(* Logix 5000 project; controller R400_500_XLS vendor 1 type 14 code 216 rev 31.11; software revision 31.01; part 31 of 32 *)
(* tags used below, declared in another part *)
   Abort1 : DINT;   // Not Used
   CycExcBuffer : UDT_CYCLE;
   CycleSequence : UDT_CYCLE_SEQUENCE;
   DintBuffer : DINT[5];
   DRYING : DINT;   // Drying id number
   M : DINT[5];   // Memory Bits
   OneShot : DINT[1];
   ONS_FC64 : DINT;
   PREWASH_1 : DINT;   // Pre-wash 1 id number
   PREWASH_2 : DINT;   // Pre-wash 2 id number
   PREWASH_3 : DINT;   // Pre-wash 3 id number
   PREWASH_4 : DINT;   // Pre-wash 4 id number
   PwExcBuffer : UDT_PW;
   PWR_UP : DINT;
   rBuffer : REAL[4];
   rIn_WSH61 : REAL;
   RINSE_1 : DINT;   // Rinse 1 id number
   RINSE_2 : DINT;   // Rinse 2 id number
   RINSE_3 : DINT;   // Rinse 3 id number
   RinseExcBuffer : UDT_RINSE;
   Run : DINT;
   sOut_WSH61 : STRING;
   String : STRING[50];   // String
   Tmr : TIMER[107];
   WASH_1 : DINT;   // Wash 1 id number
   WASH_2 : DINT;   // Wash 2 id number
   WASH_3 : DINT;   // Wash 3 id number
   WASH_4 : DINT;   // Wash 4 id number
   WASH_5 : DINT;   // Wash 5 id number
   WshExcBuffer : UDT_WASH;
   ActualDay : DINT;
   Current_Screen : DINT;
   DateTime : DINT[7];
   Doors_Check : DINT;
   DoorSafetyCheck : BOOL;
   DoorSafetyCheckDay : DINT;
   DoorSafetyCheckMonth : DINT;
   DoorSafetyCheckYear : DINT;
   I_Ld_Dr_Cls_Sw : BOOL;   // Load door close
   I_Ld_Dr_Obs_Sw : BOOL;   // Load door obstruction switch
   I_Unld_Dr_Cls_Sw : BOOL;   // Unload door close
   I_Unld_Dr_Obs_Sw : BOOL;   // Unload door obstruction switch
   LastCheckNbrDays : DINT;
   Load : Doors;
   MaintainCloseLd : BOOL;
   MaintainCloseUnld : BOOL;
   MaintainOpenLd : BOOL;
   MaintainOpenUnld : BOOL;
   MaintenanceDueDays : DINT;
   msg : BOOL[512];
   Msg_DoorSteps : INT;   // Display Safety Door Test Messages
   ONS_WSH64 : SINT;
   RecallSafetyCheck : BOOL;
   Screen_Ctrl : DINT;   // PLC Screen Request
   Tpb : DINT[11];
   TpbImage : DINT[11];
   TreatmentPtr : DINT;
   Unit : Hrdwre;   // Unit Configuration
   UnLoad : Doors;
(* MainProgram, continued *)

ROUTINE WSH_61_Real_to_String   (* ladder *)
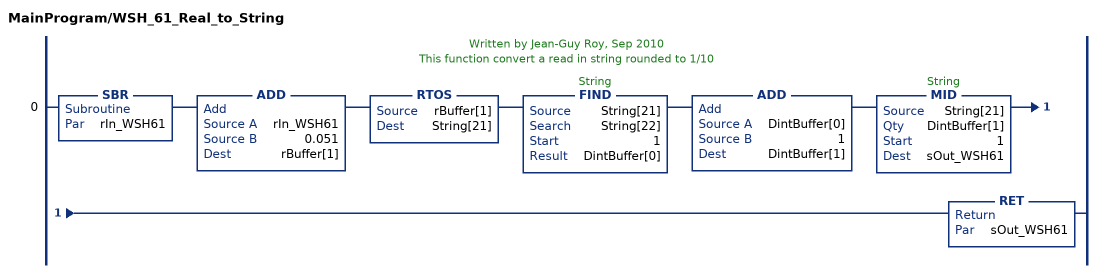
   // Written by Jean-Guy Roy, Sep 2010
   // This function convert a read in string rounded to 1/10
   0: SBR(rIn_WSH61)ADD(rIn_WSH61,0.051,rBuffer[1])RTOS(rBuffer[1],String[21])FIND(String[21],String[22],1,DintBuffer[0])ADD(DintBuffer[0],1,DintBuffer[1])MID(String[21],DintBuffer[1],1,sOut_WSH61)RET(sOut_WSH61);
END_ROUTINE

ROUTINE WSH_64_DOOR_MAINTENANCE   (* ladder *)
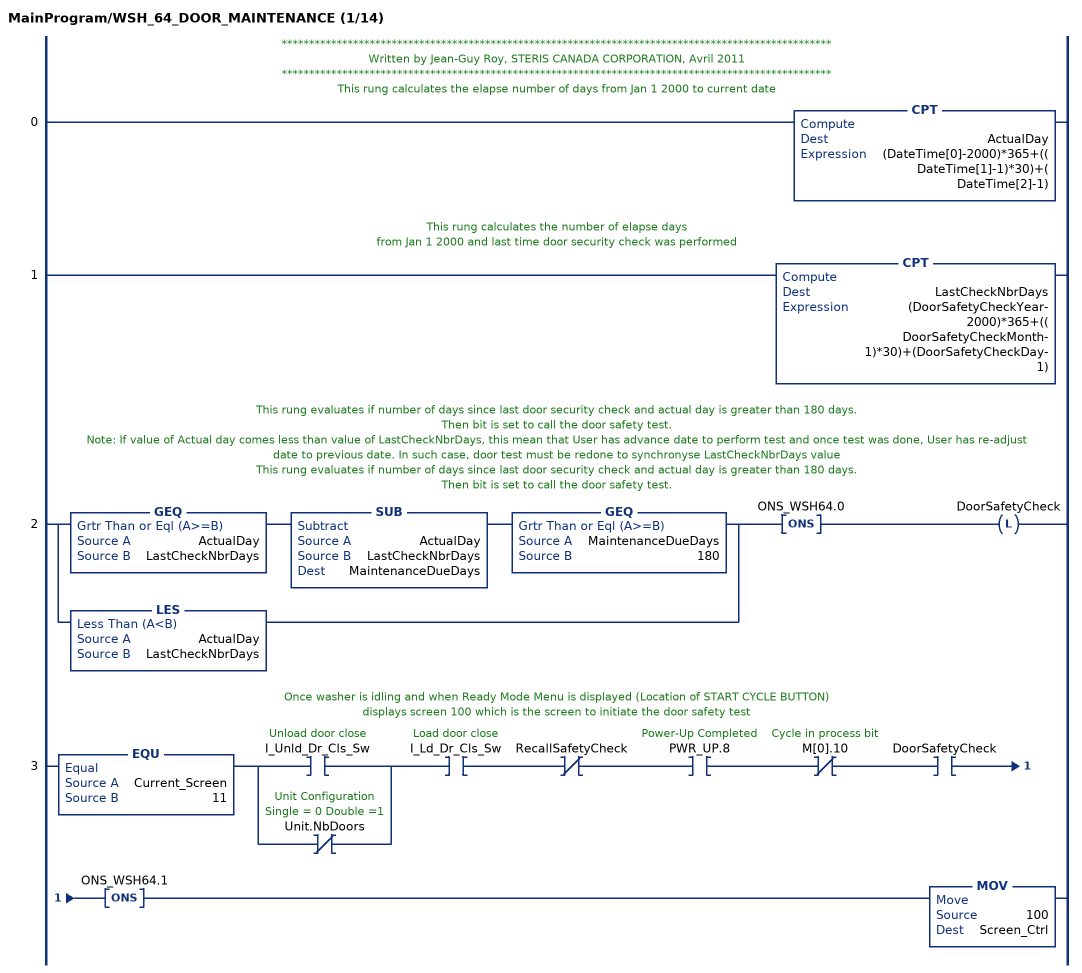
   // ****************************************************************************************************
   // Written by Jean-Guy Roy, STERIS CANADA CORPORATION, Avril 2011
   // ****************************************************************************************************
   // This rung calculates the elapse number of days from Jan 1 2000 to current date
   0: CPT(ActualDay,(DateTime[0]-2000)*365+((DateTime[1]-1)*30)+(DateTime[2]-1));
   // This rung calculates the number of elapse days
   // from Jan 1 2000 and last time door security check was performed
   1: CPT(LastCheckNbrDays,(DoorSafetyCheckYear-2000)*365+((DoorSafetyCheckMonth-1)*30)+(DoorSafetyCheckDay-1));
   // This rung evaluates if number of days since last door security check and actual day is greater than 180 days.
   // Then bit is set to call the door safety test.
   // Note: If value of Actual day comes less than value of LastCheckNbrDays, this mean that User has advance date to perform test and once test was done, User has re-adjust date to previous date. In such case, door test must be redone to synchronyse LastCheckNbrDays value
   // This rung evaluates if number of days since last door security check and actual day is greater than 180 days.
   // Then bit is set to call the door safety test.
   2: [GEQ(ActualDay,LastCheckNbrDays) SUB(ActualDay,LastCheckNbrDays,MaintenanceDueDays) GEQ(MaintenanceDueDays,180) ,LES(ActualDay,LastCheckNbrDays) ]ONS(ONS_WSH64.0)OTL(DoorSafetyCheck);
   // Once washer is idling and when Ready Mode Menu is displayed (Location of START CYCLE BUTTON)
   // displays screen 100 which is the screen to initiate the door safety test
   3: EQU(Current_Screen,11)[XIC(I_Unld_Dr_Cls_Sw) ,XIO(Unit.NbDoors) ]XIC(I_Ld_Dr_Cls_Sw)XIO(RecallSafetyCheck)XIC(PWR_UP.8)XIO(M[0].10)XIC(DoorSafetyCheck)ONS(ONS_WSH64.1)MOV(100,Screen_Ctrl);
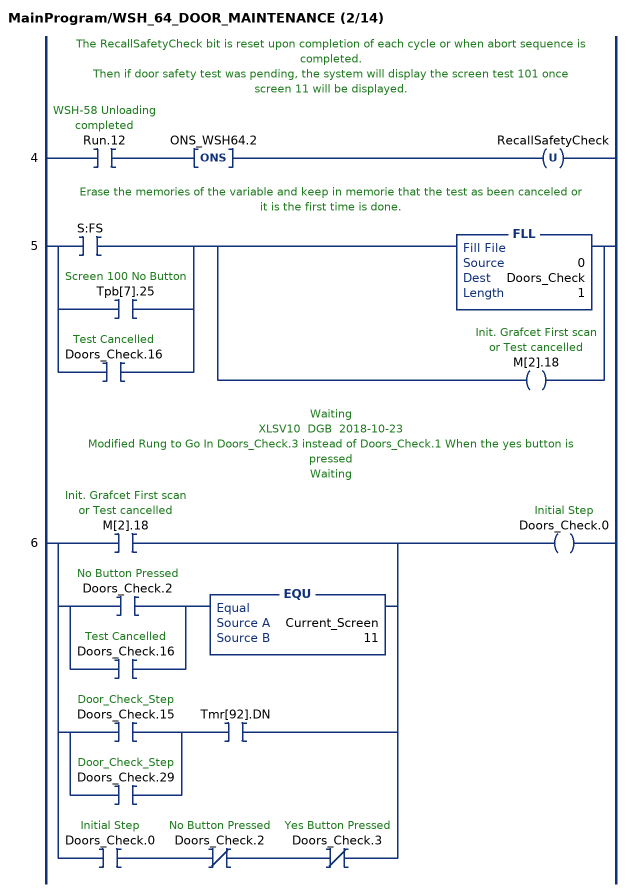
   // The RecallSafetyCheck bit is reset upon completion of each cycle or when abort sequence is completed.
   // Then if door safety test was pending, the system will display the screen test 101 once screen 11 will be displayed.
   4: XIC(Run.12)ONS(ONS_WSH64.2)OTU(RecallSafetyCheck);
   // Erase the memories of the variable and keep in memorie that the test as been canceled or it is the first time is done.
   5: [XIC(S:FS) ,XIC(Tpb[7].25) ,XIC(Doors_Check.16) ][FLL(0,Doors_Check,1) ,OTE(M[2].18) ];
   // Waiting
   // XLSV10  DGB  2018-10-23
   // Modified Rung to Go In Doors_Check.3 instead of Doors_Check.1 When the yes button is pressed
   // Waiting
   6: [XIC(M[2].18) ,[XIC(Doors_Check.2) ,XIC(Doors_Check.16) ] EQU(Current_Screen,11) ,[XIC(Doors_Check.15) ,XIC(Doors_Check.29) ] XIC(Tmr[92].DN) ,XIC(Doors_Check.0) XIO(Doors_Check.2) XIO(Doors_Check.3) ]OTE(Doors_Check.0);
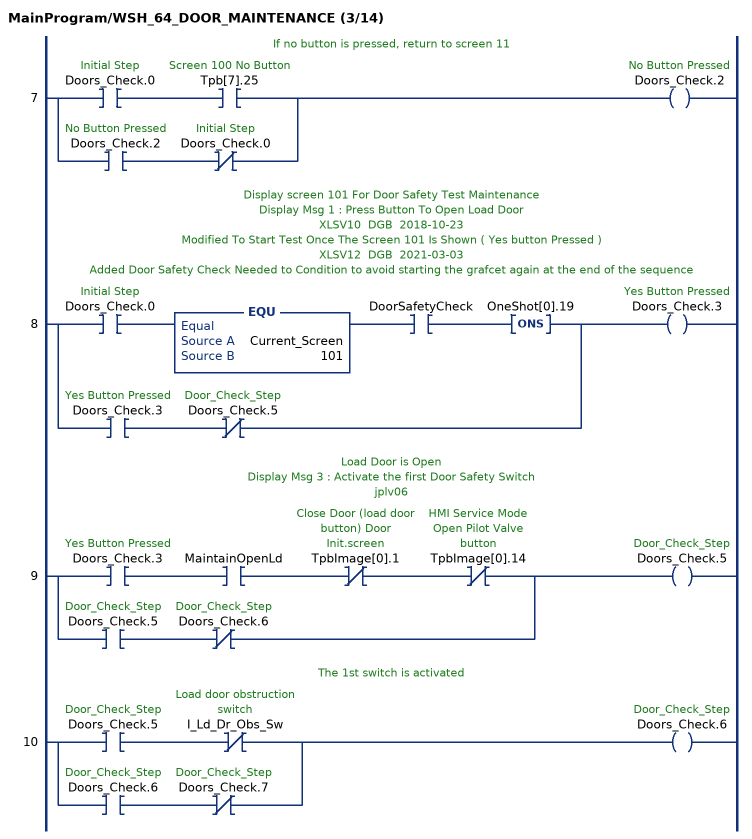
   // If no button is pressed, return to screen 11
   7: [XIC(Doors_Check.0) XIC(Tpb[7].25) ,XIC(Doors_Check.2) XIO(Doors_Check.0) ]OTE(Doors_Check.2);
   // Display screen 101 For Door Safety Test Maintenance
   // Display Msg 1 : Press Button To Open Load Door
   // XLSV10  DGB  2018-10-23
   // Modified To Start Test Once The Screen 101 Is Shown ( Yes button Pressed )
   // XLSV12  DGB  2021-03-03
   // Added Door Safety Check Needed to Condition to avoid starting the grafcet again at the end of the sequence
   8: [XIC(Doors_Check.0) EQU(Current_Screen,101) XIC(DoorSafetyCheck) ONS(OneShot[0].19) ,XIC(Doors_Check.3) XIO(Doors_Check.5) ]OTE(Doors_Check.3);
   // Load Door is Open
   // Display Msg 3 : Activate the first Door Safety Switch
   // jplv06
   9: [XIC(Doors_Check.3) XIC(MaintainOpenLd) XIO(TpbImage[0].1) XIO(TpbImage[0].14) ,XIC(Doors_Check.5) XIO(Doors_Check.6) ]OTE(Doors_Check.5);
   // The 1st switch is activated
   10: [XIC(Doors_Check.5) XIO(I_Ld_Dr_Obs_Sw) ,XIC(Doors_Check.6) XIO(Doors_Check.7) ]OTE(Doors_Check.6);
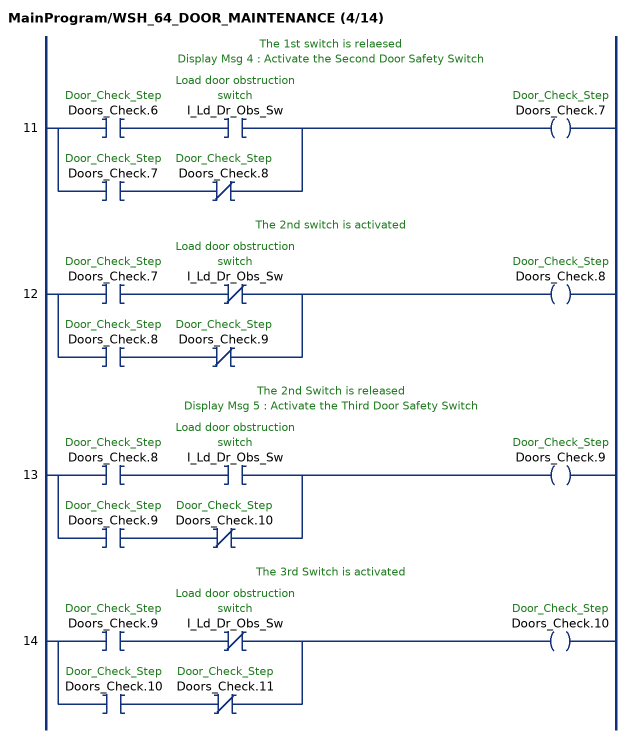
   // The 1st switch is relaesed
   // Display Msg 4 : Activate the Second Door Safety Switch
   11: [XIC(Doors_Check.6) XIC(I_Ld_Dr_Obs_Sw) ,XIC(Doors_Check.7) XIO(Doors_Check.8) ]OTE(Doors_Check.7);
   // The 2nd switch is activated
   12: [XIC(Doors_Check.7) XIO(I_Ld_Dr_Obs_Sw) ,XIC(Doors_Check.8) XIO(Doors_Check.9) ]OTE(Doors_Check.8);
   // The 2nd Switch is released
   // Display Msg 5 : Activate the Third Door Safety Switch
   13: [XIC(Doors_Check.8) XIC(I_Ld_Dr_Obs_Sw) ,XIC(Doors_Check.9) XIO(Doors_Check.10) ]OTE(Doors_Check.9);
   // The 3rd Switch is activated
   14: [XIC(Doors_Check.9) XIO(I_Ld_Dr_Obs_Sw) ,XIC(Doors_Check.10) XIO(Doors_Check.11) ]OTE(Doors_Check.10);
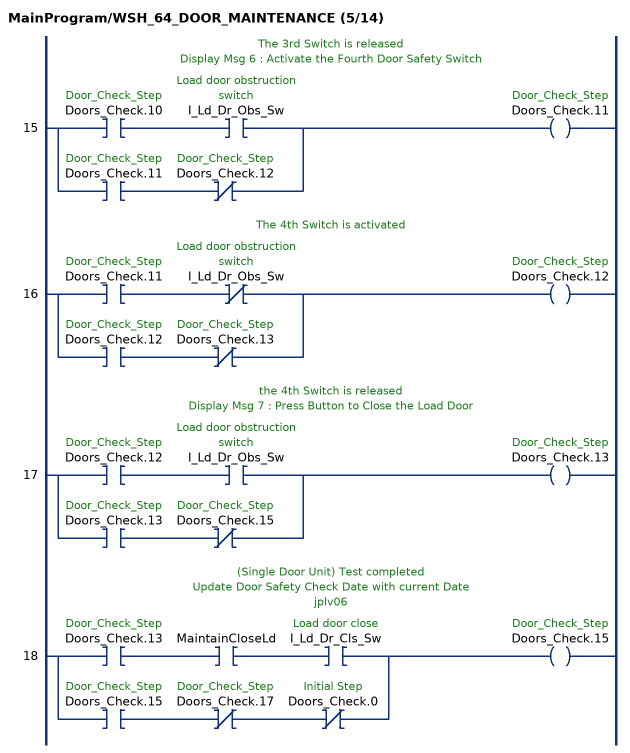
   // The 3rd Switch is released
   // Display Msg 6 : Activate the Fourth Door Safety Switch
   15: [XIC(Doors_Check.10) XIC(I_Ld_Dr_Obs_Sw) ,XIC(Doors_Check.11) XIO(Doors_Check.12) ]OTE(Doors_Check.11);
   // The 4th Switch is activated
   16: [XIC(Doors_Check.11) XIO(I_Ld_Dr_Obs_Sw) ,XIC(Doors_Check.12) XIO(Doors_Check.13) ]OTE(Doors_Check.12);
   // the 4th Switch is released
   // Display Msg 7 : Press Button to Close the Load Door
   17: [XIC(Doors_Check.12) XIC(I_Ld_Dr_Obs_Sw) ,XIC(Doors_Check.13) XIO(Doors_Check.15) ]OTE(Doors_Check.13);
   // (Single Door Unit) Test completed
   // Update Door Safety Check Date with current Date
   // jplv06
   18: [XIC(Doors_Check.13) XIC(MaintainCloseLd) XIC(I_Ld_Dr_Cls_Sw) ,XIC(Doors_Check.15) XIO(Doors_Check.17) XIO(Doors_Check.0) ]OTE(Doors_Check.15);
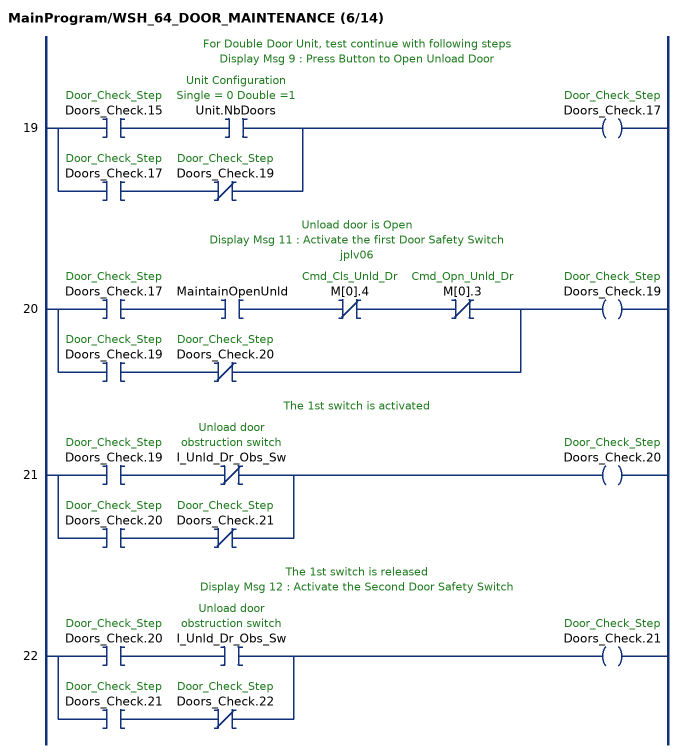
   // For Double Door Unit, test continue with following steps
   // Display Msg 9 : Press Button to Open Unload Door
   19: [XIC(Doors_Check.15) XIC(Unit.NbDoors) ,XIC(Doors_Check.17) XIO(Doors_Check.19) ]OTE(Doors_Check.17);
   // Unload door is Open
   // Display Msg 11 : Activate the first Door Safety Switch
   // jplv06
   20: [XIC(Doors_Check.17) XIC(MaintainOpenUnld) XIO(M[0].4) XIO(M[0].3) ,XIC(Doors_Check.19) XIO(Doors_Check.20) ]OTE(Doors_Check.19);
   // The 1st switch is activated
   21: [XIC(Doors_Check.19) XIO(I_Unld_Dr_Obs_Sw) ,XIC(Doors_Check.20) XIO(Doors_Check.21) ]OTE(Doors_Check.20);
   // The 1st switch is released
   // Display Msg 12 : Activate the Second Door Safety Switch
   22: [XIC(Doors_Check.20) XIC(I_Unld_Dr_Obs_Sw) ,XIC(Doors_Check.21) XIO(Doors_Check.22) ]OTE(Doors_Check.21);
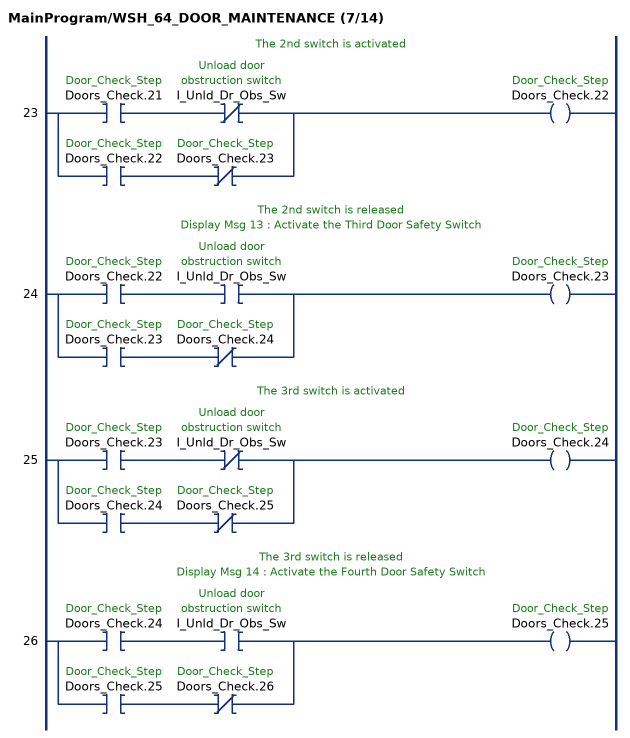
   // The 2nd switch is activated
   23: [XIC(Doors_Check.21) XIO(I_Unld_Dr_Obs_Sw) ,XIC(Doors_Check.22) XIO(Doors_Check.23) ]OTE(Doors_Check.22);
   // The 2nd switch is released
   // Display Msg 13 : Activate the Third Door Safety Switch
   24: [XIC(Doors_Check.22) XIC(I_Unld_Dr_Obs_Sw) ,XIC(Doors_Check.23) XIO(Doors_Check.24) ]OTE(Doors_Check.23);
   // The 3rd switch is activated
   25: [XIC(Doors_Check.23) XIO(I_Unld_Dr_Obs_Sw) ,XIC(Doors_Check.24) XIO(Doors_Check.25) ]OTE(Doors_Check.24);
   // The 3rd switch is released
   // Display Msg 14 : Activate the Fourth Door Safety Switch
   26: [XIC(Doors_Check.24) XIC(I_Unld_Dr_Obs_Sw) ,XIC(Doors_Check.25) XIO(Doors_Check.26) ]OTE(Doors_Check.25);
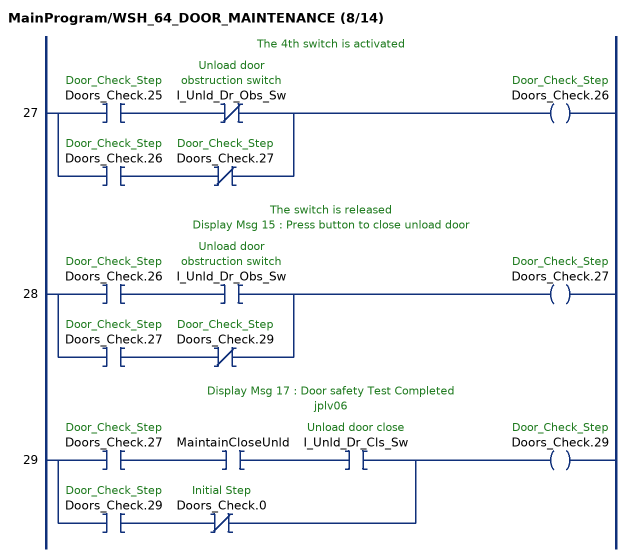
   // The 4th switch is activated
   27: [XIC(Doors_Check.25) XIO(I_Unld_Dr_Obs_Sw) ,XIC(Doors_Check.26) XIO(Doors_Check.27) ]OTE(Doors_Check.26);
   // The switch is released
   // Display Msg 15 : Press button to close unload door
   28: [XIC(Doors_Check.26) XIC(I_Unld_Dr_Obs_Sw) ,XIC(Doors_Check.27) XIO(Doors_Check.29) ]OTE(Doors_Check.27);
   // Display Msg 17 : Door safety Test Completed
   // jplv06
   29: [XIC(Doors_Check.27) XIC(MaintainCloseUnld) XIC(I_Unld_Dr_Cls_Sw) ,XIC(Doors_Check.29) XIO(Doors_Check.0) ]OTE(Doors_Check.29);
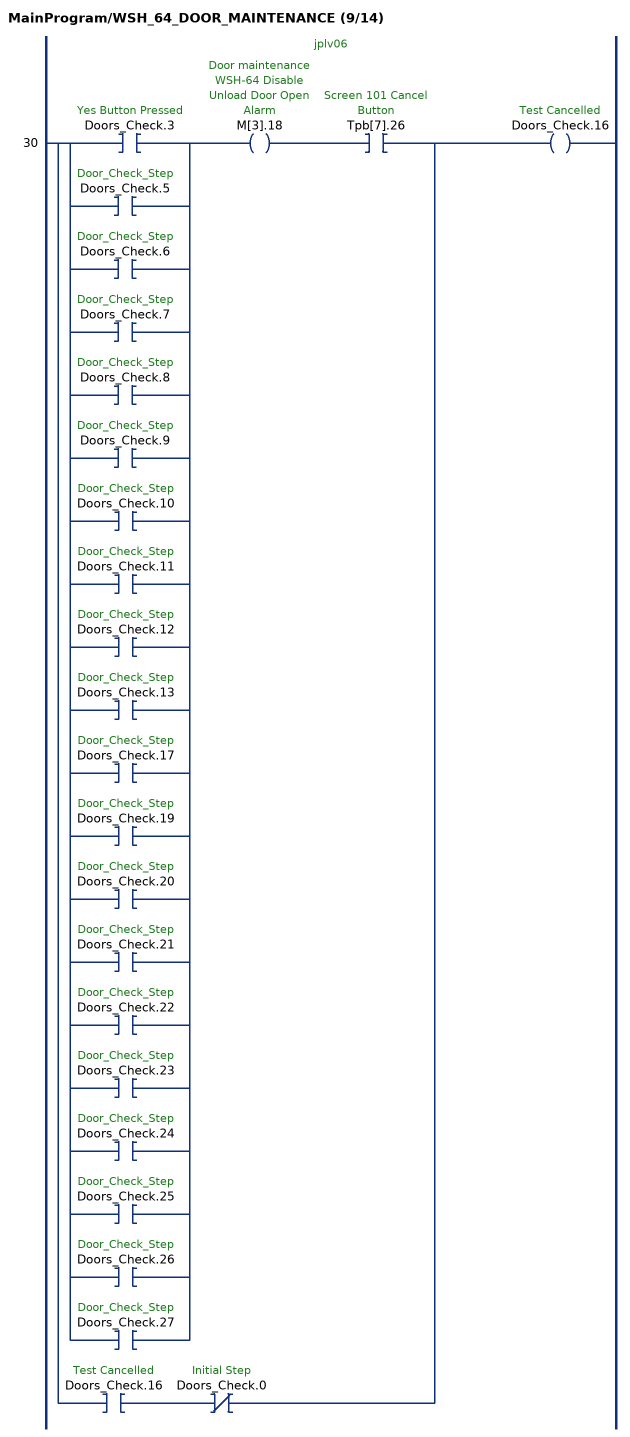
   // jplv06
   30: [[XIC(Doors_Check.3) ,XIC(Doors_Check.5) ,XIC(Doors_Check.6) ,XIC(Doors_Check.7) ,XIC(Doors_Check.8) ,XIC(Doors_Check.9) ,XIC(Doors_Check.10) ,XIC(Doors_Check.11) ,XIC(Doors_Check.12) ,XIC(Doors_Check.13) ,XIC(Doors_Check.17) ,XIC(Doors_Check.19) ,XIC(Doors_Check.20) ,XIC(Doors_Check.21) ,XIC(Doors_Check.22) ,XIC(Doors_Check.23) ,XIC(Doors_Check.24) ,XIC(Doors_Check.25) ,XIC(Doors_Check.26) ,XIC(Doors_Check.27) ] OTE(M[3].18) XIC(Tpb[7].26) ,XIC(Doors_Check.16) XIO(Doors_Check.0) ]OTE(Doors_Check.16);
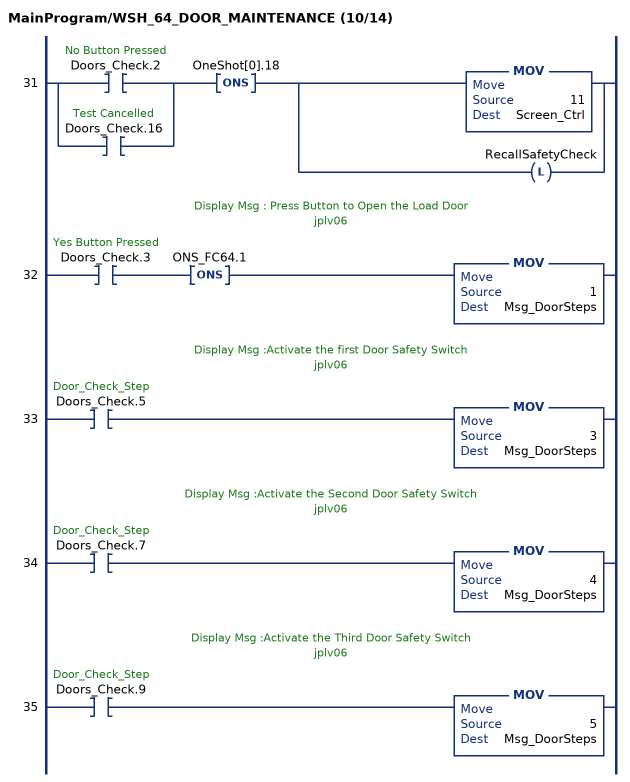
   31: [XIC(Doors_Check.2) ,XIC(Doors_Check.16) ]ONS(OneShot[0].18)[MOV(11,Screen_Ctrl) ,OTL(RecallSafetyCheck) ];
   // Display Msg : Press Button to Open the Load Door
   // jplv06
   32: XIC(Doors_Check.3)ONS(ONS_FC64.1)MOV(1,Msg_DoorSteps);
   // Display Msg :Activate the first Door Safety Switch
   // jplv06
   33: XIC(Doors_Check.5)MOV(3,Msg_DoorSteps);
   // Display Msg :Activate the Second Door Safety Switch
   // jplv06
   34: XIC(Doors_Check.7)MOV(4,Msg_DoorSteps);
   // Display Msg :Activate the Third Door Safety Switch
   // jplv06
   35: XIC(Doors_Check.9)MOV(5,Msg_DoorSteps);
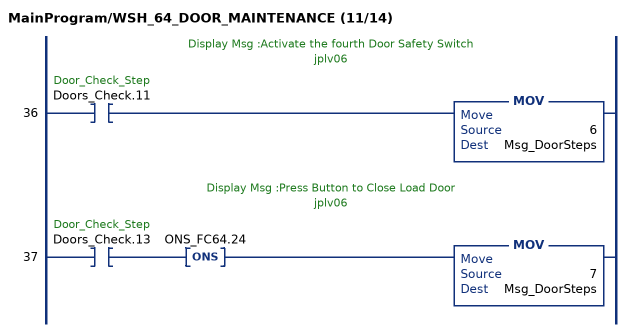
   // Display Msg :Activate the fourth Door Safety Switch
   // jplv06
   36: XIC(Doors_Check.11)MOV(6,Msg_DoorSteps);
   // Display Msg :Press Button to Close Load Door
   // jplv06
   37: XIC(Doors_Check.13)ONS(ONS_FC64.24)MOV(7,Msg_DoorSteps);
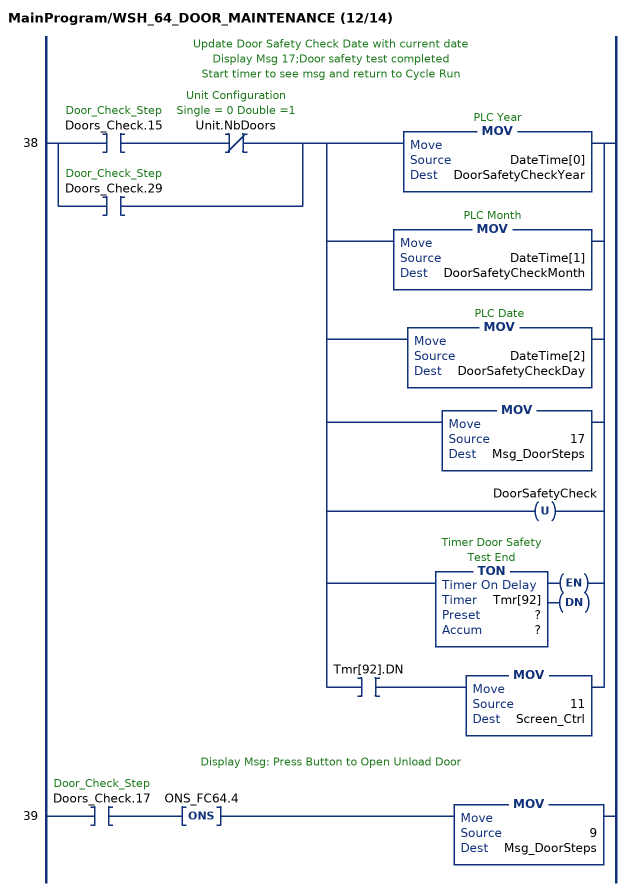
   // Update Door Safety Check Date with current date
   // Display Msg 17;Door safety test completed
   // Start timer to see msg and return to Cycle Run
   38: [XIC(Doors_Check.15) XIO(Unit.NbDoors) ,XIC(Doors_Check.29) ][MOV(DateTime[0],DoorSafetyCheckYear) ,MOV(DateTime[1],DoorSafetyCheckMonth) ,MOV(DateTime[2],DoorSafetyCheckDay) ,MOV(17,Msg_DoorSteps) ,OTU(DoorSafetyCheck) ,TON(Tmr[92],?,?) ,XIC(Tmr[92].DN) MOV(11,Screen_Ctrl) ];
   // Display Msg: Press Button to Open Unload Door
   39: XIC(Doors_Check.17)ONS(ONS_FC64.4)MOV(9,Msg_DoorSteps);
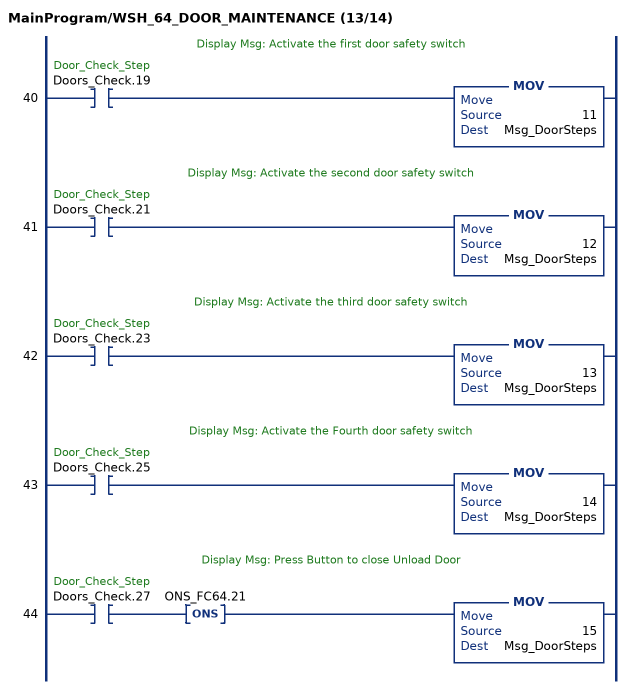
   // Display Msg: Activate the first door safety switch
   40: XIC(Doors_Check.19)MOV(11,Msg_DoorSteps);
   // Display Msg: Activate the second door safety switch
   41: XIC(Doors_Check.21)MOV(12,Msg_DoorSteps);
   // Display Msg: Activate the third door safety switch
   42: XIC(Doors_Check.23)MOV(13,Msg_DoorSteps);
   // Display Msg: Activate the Fourth door safety switch
   43: XIC(Doors_Check.25)MOV(14,Msg_DoorSteps);
   // Display Msg: Press Button to close Unload Door
   44: XIC(Doors_Check.27)ONS(ONS_FC64.21)MOV(15,Msg_DoorSteps);
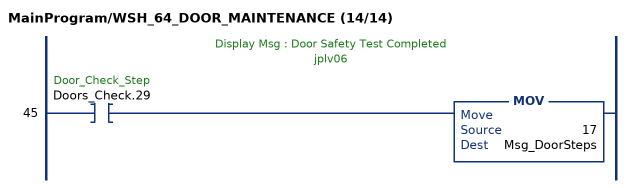
   // Display Msg : Door Safety Test Completed
   // jplv06
   45: XIC(Doors_Check.29)MOV(17,Msg_DoorSteps);
END_ROUTINE

ROUTINE WSH_8_PERFOM_CYCLE   (* ladder *)
// Cycle function to
// Process Recirculated Treatment, Final Rinse Treatment and Drying Treatment.
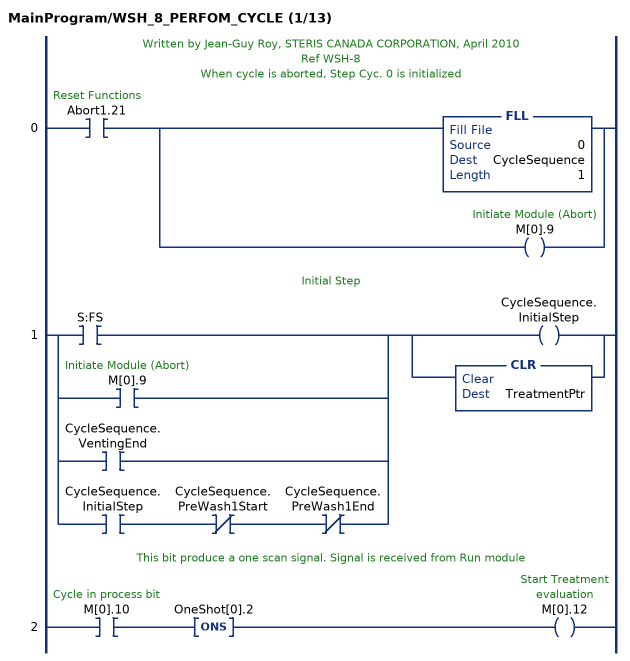
   // Written by Jean-Guy Roy, STERIS CANADA CORPORATION, April 2010
   // Ref WSH-8
   // When cycle is aborted, Step Cyc. 0 is initialized
   0: XIC(Abort1.21)[FLL(0,CycleSequence,1) ,OTE(M[0].9) ];
   // Initial Step
   1: [XIC(S:FS) ,XIC(M[0].9) ,XIC(CycleSequence.VentingEnd) ,XIC(CycleSequence.InitialStep) XIO(CycleSequence.PreWash1Start) XIO(CycleSequence.PreWash1End) ][OTE(CycleSequence.InitialStep) ,CLR(TreatmentPtr) ];
   // This bit produce a one scan signal. Signal is received from Run module
   2: XIC(M[0].10)ONS(OneShot[0].2)OTE(M[0].12);
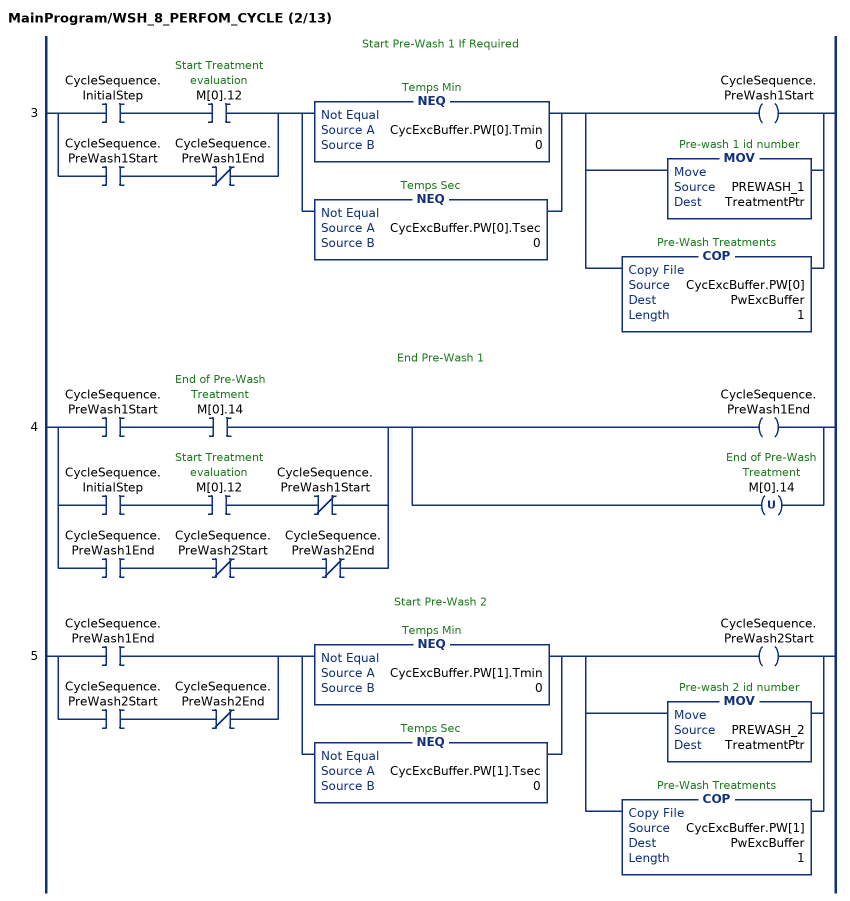
   // Start Pre-Wash 1 If Required
   3: [XIC(CycleSequence.InitialStep) XIC(M[0].12) ,XIC(CycleSequence.PreWash1Start) XIO(CycleSequence.PreWash1End) ][NEQ(CycExcBuffer.PW[0].Tmin,0) ,NEQ(CycExcBuffer.PW[0].Tsec,0) ][OTE(CycleSequence.PreWash1Start) ,MOV(PREWASH_1,TreatmentPtr) ,COP(CycExcBuffer.PW[0],PwExcBuffer,1) ];
   // End Pre-Wash 1
   4: [XIC(CycleSequence.PreWash1Start) XIC(M[0].14) ,XIC(CycleSequence.InitialStep) XIC(M[0].12) XIO(CycleSequence.PreWash1Start) ,XIC(CycleSequence.PreWash1End) XIO(CycleSequence.PreWash2Start) XIO(CycleSequence.PreWash2End) ][OTE(CycleSequence.PreWash1End) ,OTU(M[0].14) ];
   // Start Pre-Wash 2
   5: [XIC(CycleSequence.PreWash1End) ,XIC(CycleSequence.PreWash2Start) XIO(CycleSequence.PreWash2End) ][NEQ(CycExcBuffer.PW[1].Tmin,0) ,NEQ(CycExcBuffer.PW[1].Tsec,0) ][OTE(CycleSequence.PreWash2Start) ,MOV(PREWASH_2,TreatmentPtr) ,COP(CycExcBuffer.PW[1],PwExcBuffer,1) ];
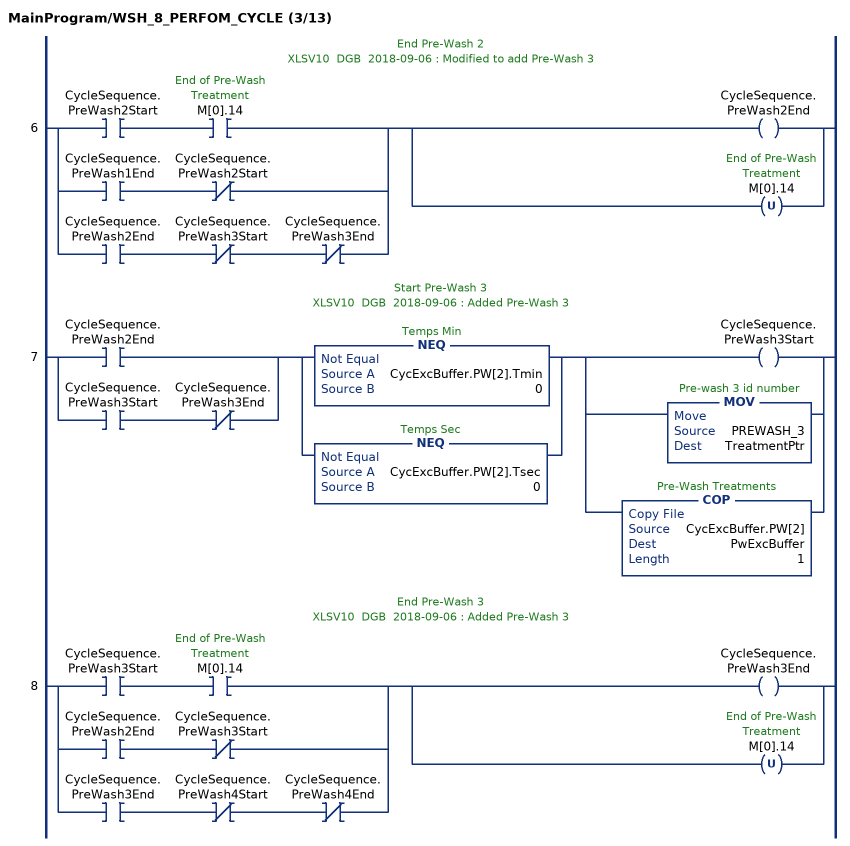
   // End Pre-Wash 2
   // XLSV10  DGB  2018-09-06 : Modified to add Pre-Wash 3
   6: [XIC(CycleSequence.PreWash2Start) XIC(M[0].14) ,XIC(CycleSequence.PreWash1End) XIO(CycleSequence.PreWash2Start) ,XIC(CycleSequence.PreWash2End) XIO(CycleSequence.PreWash3Start) XIO(CycleSequence.PreWash3End) ][OTE(CycleSequence.PreWash2End) ,OTU(M[0].14) ];
   // Start Pre-Wash 3
   // XLSV10  DGB  2018-09-06 : Added Pre-Wash 3
   7: [XIC(CycleSequence.PreWash2End) ,XIC(CycleSequence.PreWash3Start) XIO(CycleSequence.PreWash3End) ][NEQ(CycExcBuffer.PW[2].Tmin,0) ,NEQ(CycExcBuffer.PW[2].Tsec,0) ][OTE(CycleSequence.PreWash3Start) ,MOV(PREWASH_3,TreatmentPtr) ,COP(CycExcBuffer.PW[2],PwExcBuffer,1) ];
   // End Pre-Wash 3
   // XLSV10  DGB  2018-09-06 : Added Pre-Wash 3
   8: [XIC(CycleSequence.PreWash3Start) XIC(M[0].14) ,XIC(CycleSequence.PreWash2End) XIO(CycleSequence.PreWash3Start) ,XIC(CycleSequence.PreWash3End) XIO(CycleSequence.PreWash4Start) XIO(CycleSequence.PreWash4End) ][OTE(CycleSequence.PreWash3End) ,OTU(M[0].14) ];
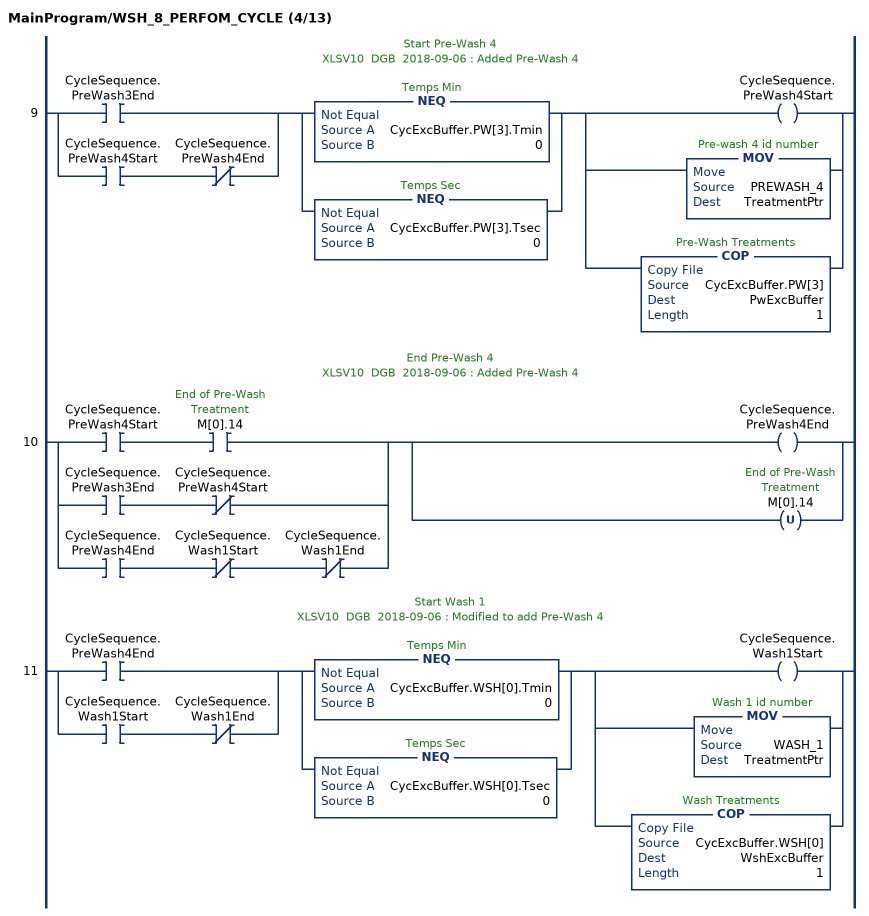
   // Start Pre-Wash 4
   // XLSV10  DGB  2018-09-06 : Added Pre-Wash 4
   9: [XIC(CycleSequence.PreWash3End) ,XIC(CycleSequence.PreWash4Start) XIO(CycleSequence.PreWash4End) ][NEQ(CycExcBuffer.PW[3].Tmin,0) ,NEQ(CycExcBuffer.PW[3].Tsec,0) ][OTE(CycleSequence.PreWash4Start) ,MOV(PREWASH_4,TreatmentPtr) ,COP(CycExcBuffer.PW[3],PwExcBuffer,1) ];
   // End Pre-Wash 4
   // XLSV10  DGB  2018-09-06 : Added Pre-Wash 4
   10: [XIC(CycleSequence.PreWash4Start) XIC(M[0].14) ,XIC(CycleSequence.PreWash3End) XIO(CycleSequence.PreWash4Start) ,XIC(CycleSequence.PreWash4End) XIO(CycleSequence.Wash1Start) XIO(CycleSequence.Wash1End) ][OTE(CycleSequence.PreWash4End) ,OTU(M[0].14) ];
   // Start Wash 1
   // XLSV10  DGB  2018-09-06 : Modified to add Pre-Wash 4
   11: [XIC(CycleSequence.PreWash4End) ,XIC(CycleSequence.Wash1Start) XIO(CycleSequence.Wash1End) ][NEQ(CycExcBuffer.WSH[0].Tmin,0) ,NEQ(CycExcBuffer.WSH[0].Tsec,0) ][OTE(CycleSequence.Wash1Start) ,MOV(WASH_1,TreatmentPtr) ,COP(CycExcBuffer.WSH[0],WshExcBuffer,1) ];
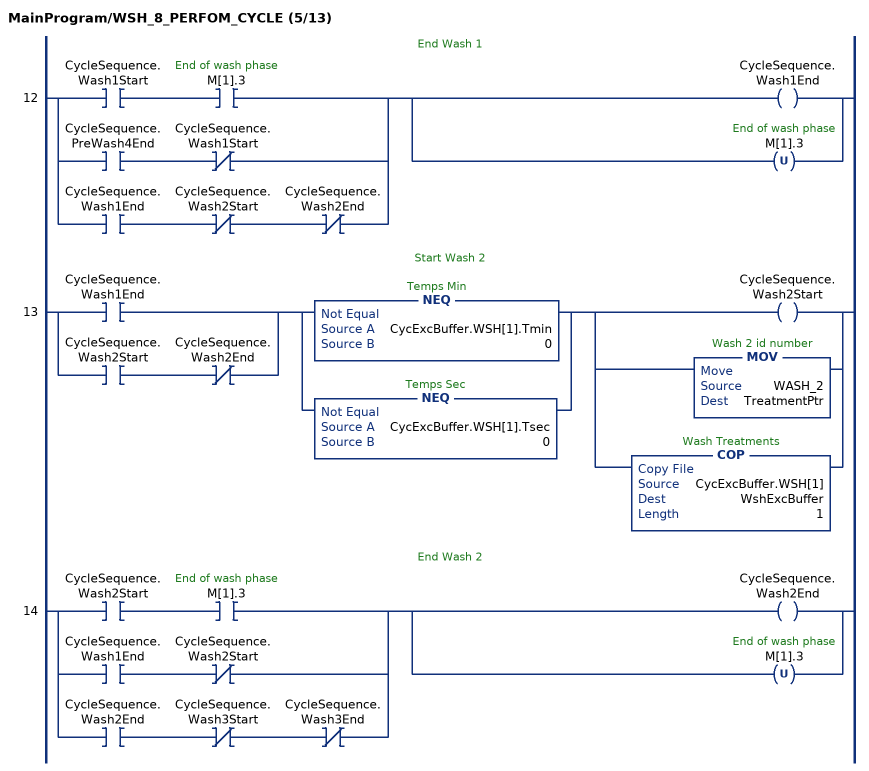
   // End Wash 1
   12: [XIC(CycleSequence.Wash1Start) XIC(M[1].3) ,XIC(CycleSequence.PreWash4End) XIO(CycleSequence.Wash1Start) ,XIC(CycleSequence.Wash1End) XIO(CycleSequence.Wash2Start) XIO(CycleSequence.Wash2End) ][OTE(CycleSequence.Wash1End) ,OTU(M[1].3) ];
   // Start Wash 2
   13: [XIC(CycleSequence.Wash1End) ,XIC(CycleSequence.Wash2Start) XIO(CycleSequence.Wash2End) ][NEQ(CycExcBuffer.WSH[1].Tmin,0) ,NEQ(CycExcBuffer.WSH[1].Tsec,0) ][OTE(CycleSequence.Wash2Start) ,MOV(WASH_2,TreatmentPtr) ,COP(CycExcBuffer.WSH[1],WshExcBuffer,1) ];
   // End Wash 2
   14: [XIC(CycleSequence.Wash2Start) XIC(M[1].3) ,XIC(CycleSequence.Wash1End) XIO(CycleSequence.Wash2Start) ,XIC(CycleSequence.Wash2End) XIO(CycleSequence.Wash3Start) XIO(CycleSequence.Wash3End) ][OTE(CycleSequence.Wash2End) ,OTU(M[1].3) ];
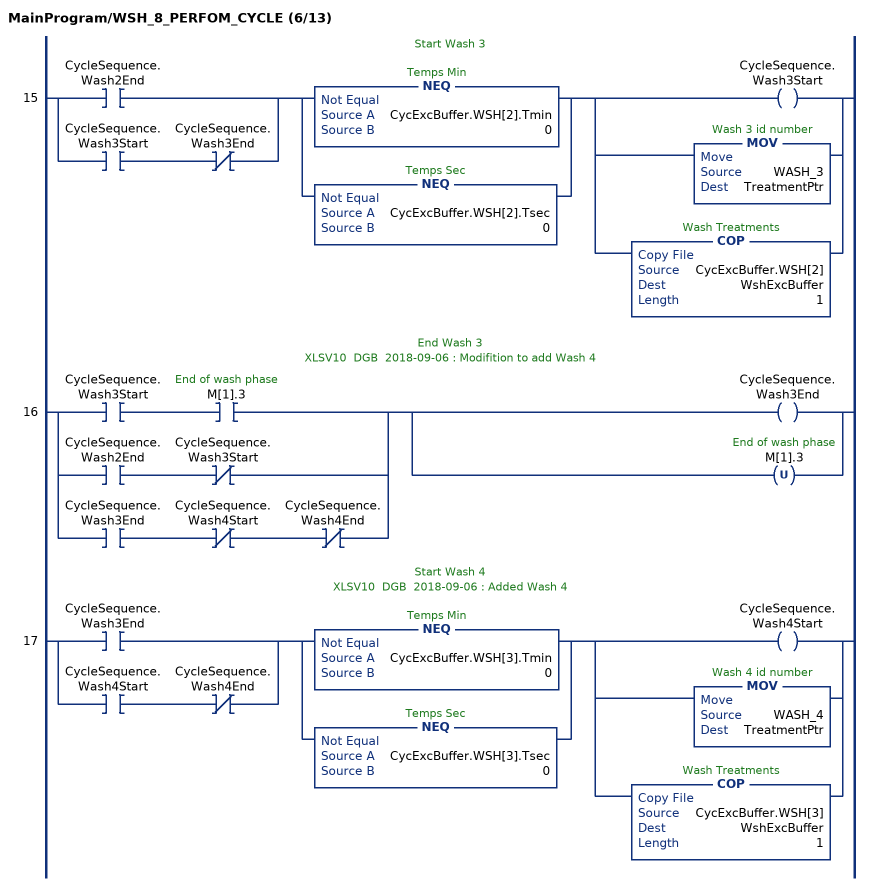
   // Start Wash 3
   15: [XIC(CycleSequence.Wash2End) ,XIC(CycleSequence.Wash3Start) XIO(CycleSequence.Wash3End) ][NEQ(CycExcBuffer.WSH[2].Tmin,0) ,NEQ(CycExcBuffer.WSH[2].Tsec,0) ][OTE(CycleSequence.Wash3Start) ,MOV(WASH_3,TreatmentPtr) ,COP(CycExcBuffer.WSH[2],WshExcBuffer,1) ];
   // End Wash 3
   // XLSV10  DGB  2018-09-06 : Modifition to add Wash 4
   16: [XIC(CycleSequence.Wash3Start) XIC(M[1].3) ,XIC(CycleSequence.Wash2End) XIO(CycleSequence.Wash3Start) ,XIC(CycleSequence.Wash3End) XIO(CycleSequence.Wash4Start) XIO(CycleSequence.Wash4End) ][OTE(CycleSequence.Wash3End) ,OTU(M[1].3) ];
   // Start Wash 4
   // XLSV10  DGB  2018-09-06 : Added Wash 4
   17: [XIC(CycleSequence.Wash3End) ,XIC(CycleSequence.Wash4Start) XIO(CycleSequence.Wash4End) ][NEQ(CycExcBuffer.WSH[3].Tmin,0) ,NEQ(CycExcBuffer.WSH[3].Tsec,0) ][OTE(CycleSequence.Wash4Start) ,MOV(WASH_4,TreatmentPtr) ,COP(CycExcBuffer.WSH[3],WshExcBuffer,1) ];
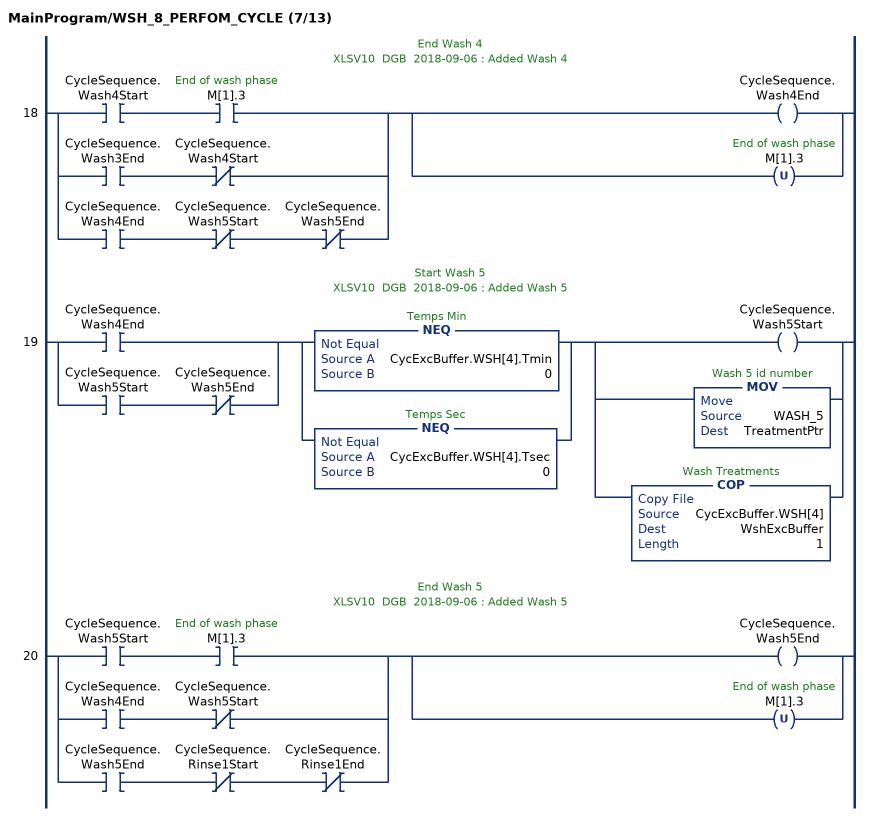
   // End Wash 4
   // XLSV10  DGB  2018-09-06 : Added Wash 4
   18: [XIC(CycleSequence.Wash4Start) XIC(M[1].3) ,XIC(CycleSequence.Wash3End) XIO(CycleSequence.Wash4Start) ,XIC(CycleSequence.Wash4End) XIO(CycleSequence.Wash5Start) XIO(CycleSequence.Wash5End) ][OTE(CycleSequence.Wash4End) ,OTU(M[1].3) ];
   // Start Wash 5
   // XLSV10  DGB  2018-09-06 : Added Wash 5
   19: [XIC(CycleSequence.Wash4End) ,XIC(CycleSequence.Wash5Start) XIO(CycleSequence.Wash5End) ][NEQ(CycExcBuffer.WSH[4].Tmin,0) ,NEQ(CycExcBuffer.WSH[4].Tsec,0) ][OTE(CycleSequence.Wash5Start) ,MOV(WASH_5,TreatmentPtr) ,COP(CycExcBuffer.WSH[4],WshExcBuffer,1) ];
   // End Wash 5
   // XLSV10  DGB  2018-09-06 : Added Wash 5
   20: [XIC(CycleSequence.Wash5Start) XIC(M[1].3) ,XIC(CycleSequence.Wash4End) XIO(CycleSequence.Wash5Start) ,XIC(CycleSequence.Wash5End) XIO(CycleSequence.Rinse1Start) XIO(CycleSequence.Rinse1End) ][OTE(CycleSequence.Wash5End) ,OTU(M[1].3) ];
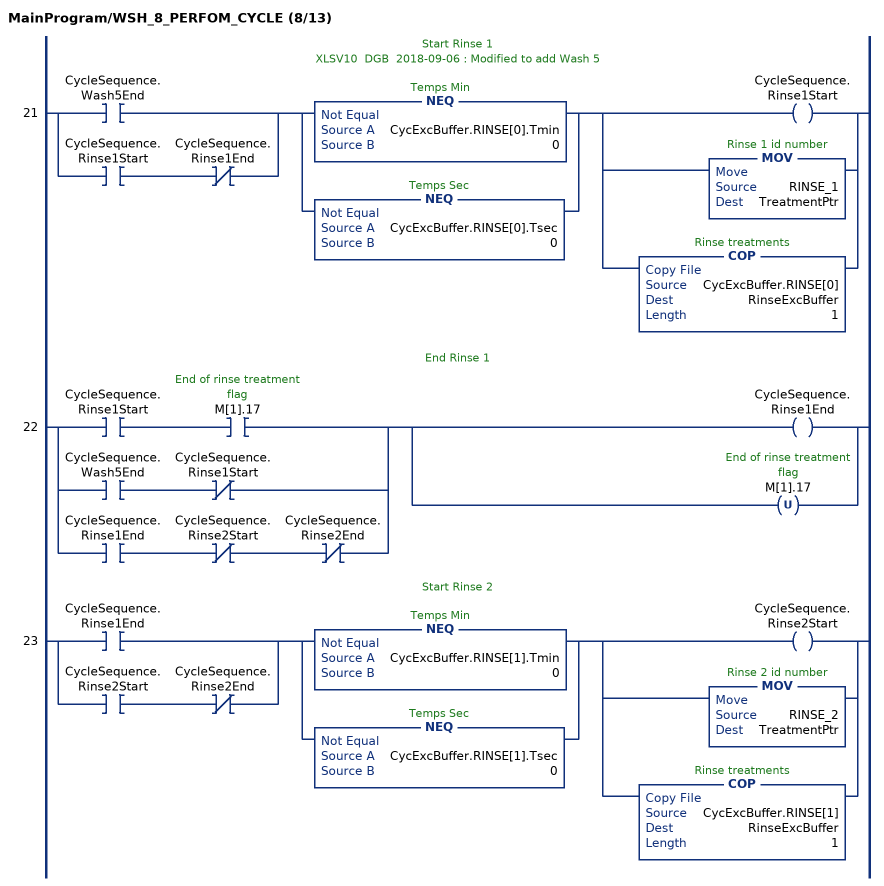
   // Start Rinse 1
   // XLSV10  DGB  2018-09-06 : Modified to add Wash 5
   21: [XIC(CycleSequence.Wash5End) ,XIC(CycleSequence.Rinse1Start) XIO(CycleSequence.Rinse1End) ][NEQ(CycExcBuffer.RINSE[0].Tmin,0) ,NEQ(CycExcBuffer.RINSE[0].Tsec,0) ][OTE(CycleSequence.Rinse1Start) ,MOV(RINSE_1,TreatmentPtr) ,COP(CycExcBuffer.RINSE[0],RinseExcBuffer,1) ];
   // End Rinse 1
   22: [XIC(CycleSequence.Rinse1Start) XIC(M[1].17) ,XIC(CycleSequence.Wash5End) XIO(CycleSequence.Rinse1Start) ,XIC(CycleSequence.Rinse1End) XIO(CycleSequence.Rinse2Start) XIO(CycleSequence.Rinse2End) ][OTE(CycleSequence.Rinse1End) ,OTU(M[1].17) ];
   // Start Rinse 2
   23: [XIC(CycleSequence.Rinse1End) ,XIC(CycleSequence.Rinse2Start) XIO(CycleSequence.Rinse2End) ][NEQ(CycExcBuffer.RINSE[1].Tmin,0) ,NEQ(CycExcBuffer.RINSE[1].Tsec,0) ][OTE(CycleSequence.Rinse2Start) ,MOV(RINSE_2,TreatmentPtr) ,COP(CycExcBuffer.RINSE[1],RinseExcBuffer,1) ];
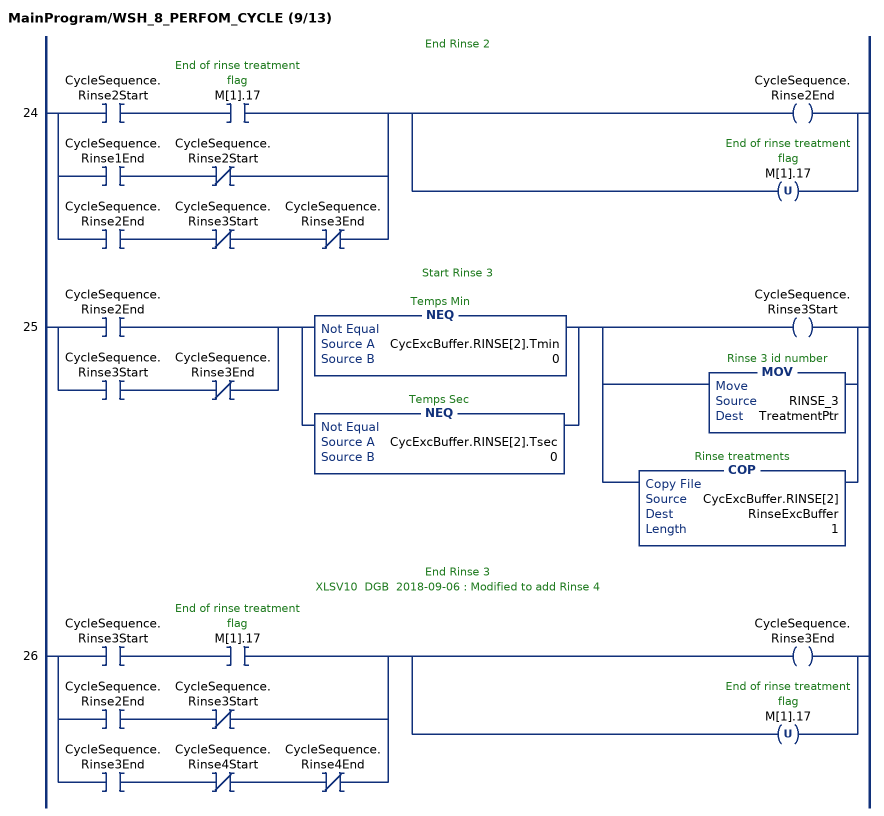
   // End Rinse 2
   24: [XIC(CycleSequence.Rinse2Start) XIC(M[1].17) ,XIC(CycleSequence.Rinse1End) XIO(CycleSequence.Rinse2Start) ,XIC(CycleSequence.Rinse2End) XIO(CycleSequence.Rinse3Start) XIO(CycleSequence.Rinse3End) ][OTE(CycleSequence.Rinse2End) ,OTU(M[1].17) ];
   // Start Rinse 3
   25: [XIC(CycleSequence.Rinse2End) ,XIC(CycleSequence.Rinse3Start) XIO(CycleSequence.Rinse3End) ][NEQ(CycExcBuffer.RINSE[2].Tmin,0) ,NEQ(CycExcBuffer.RINSE[2].Tsec,0) ][OTE(CycleSequence.Rinse3Start) ,MOV(RINSE_3,TreatmentPtr) ,COP(CycExcBuffer.RINSE[2],RinseExcBuffer,1) ];
   // End Rinse 3
   // XLSV10  DGB  2018-09-06 : Modified to add Rinse 4
   26: [XIC(CycleSequence.Rinse3Start) XIC(M[1].17) ,XIC(CycleSequence.Rinse2End) XIO(CycleSequence.Rinse3Start) ,XIC(CycleSequence.Rinse3End) XIO(CycleSequence.Rinse4Start) XIO(CycleSequence.Rinse4End) ][OTE(CycleSequence.Rinse3End) ,OTU(M[1].17) ];
